(* IEC 61131-3 sources: codesys-conveyor-sorting/src, 4 files *)

(* ---- E_ConveyorState.st ---- *)
// DUT: E_ConveyorState
// States of the conveyor sorting station.
// Numbering in steps of 10 leaves room for new states later.

{attribute 'qualified_only'}
{attribute 'strict'}
TYPE E_ConveyorState :
(
    IDLE        := 0,   // Conveyor stopped, waiting for start
    RUNNING     := 10,  // Conveyor running, waiting for a part at the infeed
    CLASSIFYING := 20,  // Part detected, reading classification sensors
    TRANSPORT   := 30,  // Part travelling to the diverter, jam timer active
    DIVERTING   := 40,  // Diverter pulse active, part counted at the end
    FAULT       := 90,  // Jam detected, conveyor stopped, waiting for reset
    ESTOP       := 99   // E-stop active, all outputs off
);
END_TYPE

(* ---- E_PartType.st ---- *)
// DUT: E_PartType
// Result of the part classification at the infeed.

{attribute 'qualified_only'}
{attribute 'strict'}
TYPE E_PartType :
(
    NONE   := 0,  // No part being tracked
    TYPE_A := 1,  // Goes to bin A
    TYPE_B := 2,  // Goes to bin B
    REJECT := 3   // Unknown part (both or neither sensor), runs to reject bin
);
END_TYPE

(* ---- GVL_IO.st ---- *)
// GVL: GVL_IO
// Inputs and outputs of the sorting station.
// In this project they are driven by the CODESYS visualisation (simulation).
// On real hardware each variable would be mapped to a physical channel
// in the I/O configuration of the fieldbus device.

{attribute 'qualified_only'}
VAR_GLOBAL
    // ---- Digital inputs ----
    xStartPB         : BOOL;          // Start push button (TRUE = pressed)
    xStopPB          : BOOL;          // Stop push button (TRUE = pressed)
    xResetPB         : BOOL;          // Fault reset push button
    xEStopOK         : BOOL := TRUE;  // E-stop circuit healthy (NC contact, TRUE = OK)
    xPartAtEntry     : BOOL;          // Photo sensor at the infeed
    xSensorTypeA     : BOOL;          // Classification sensor, TRUE = type A
    xSensorTypeB     : BOOL;          // Classification sensor, TRUE = type B
    xPartAtDiverter  : BOOL;          // Photo sensor at the diverter position

    // ---- Digital outputs ----
    xConveyorRun     : BOOL;          // Conveyor motor contactor / VFD run command
    xDiverterA       : BOOL;          // Pneumatic diverter to bin A
    xDiverterB       : BOOL;          // Pneumatic diverter to bin B
    xLampRunning     : BOOL;          // Green lamp
    xLampFault       : BOOL;          // Red lamp (steady = jam, blinking = E-stop)
END_VAR

(* ---- PLC_PRG.st ---- *)
// =====================================================================
// POU: PLC_PRG (Program, Structured Text)
// Conveyor sorting station - main state machine
//
// Sequence: IDLE -> RUNNING -> CLASSIFYING -> TRANSPORT -> DIVERTING -> RUNNING
// Faults:   jam timeout -> FAULT, E-stop -> ESTOP (both need reset, then start)
//
// Note: the real E-stop is a hardwired safety circuit. The PLC only
// monitors it (xEStopOK) to stop the sequence and show the state.
// =====================================================================

// ---------------- DECLARATION (top pane in CODESYS) ----------------
PROGRAM PLC_PRG
VAR
    eState            : E_ConveyorState := E_ConveyorState.IDLE;
    ePartType         : E_PartType := E_PartType.NONE;
    xStopRequest      : BOOL;     // Stop pressed: finish the current part, then stop

    // Edge detection
    rtStart           : R_TRIG;
    rtReset           : R_TRIG;
    rtPartAtEntry     : R_TRIG;
    rtPartAtDiverter  : R_TRIG;

    // Timers
    tonJam            : TON;      // Part must reach the diverter within T_JAM_TIMEOUT
    tonDivert         : TON;      // Length of the diverter pulse
    tonBlink          : TON;      // Blink clock for the fault lamp
    xBlink            : BOOL;

    // Production counters (read later by the OPC UA data logger)
    udiCountA         : UDINT;
    udiCountB         : UDINT;
    udiCountReject    : UDINT;
    udiCountJams      : UDINT;
END_VAR
VAR CONSTANT
    T_JAM_TIMEOUT     : TIME := T#5S;
    T_DIVERT_PULSE    : TIME := T#500MS;
    T_BLINK           : TIME := T#500MS;
END_VAR

// ---------------- IMPLEMENTATION (bottom pane in CODESYS) ----------------

// ---- Edge detection ----
rtStart(CLK := GVL_IO.xStartPB);
rtReset(CLK := GVL_IO.xResetPB);
rtPartAtEntry(CLK := GVL_IO.xPartAtEntry);
rtPartAtDiverter(CLK := GVL_IO.xPartAtDiverter);

// ---- Timers (called every scan, outside the CASE) ----
tonJam(IN := (eState = E_ConveyorState.TRANSPORT), PT := T_JAM_TIMEOUT);
tonDivert(IN := (eState = E_ConveyorState.DIVERTING), PT := T_DIVERT_PULSE);
tonBlink(IN := NOT tonBlink.Q, PT := T_BLINK);
IF tonBlink.Q THEN
    xBlink := NOT xBlink;
END_IF

// ---- E-stop has priority over every state ----
IF NOT GVL_IO.xEStopOK THEN
    eState := E_ConveyorState.ESTOP;
END_IF

// ---- Stop request is latched and handled by the states ----
IF GVL_IO.xStopPB THEN
    xStopRequest := TRUE;
END_IF

// ---- State machine ----
CASE eState OF

    E_ConveyorState.IDLE:
        xStopRequest := FALSE;
        ePartType := E_PartType.NONE;
        IF rtStart.Q AND GVL_IO.xEStopOK THEN
            eState := E_ConveyorState.RUNNING;
        END_IF

    E_ConveyorState.RUNNING:
        IF xStopRequest THEN
            eState := E_ConveyorState.IDLE;
        ELSIF rtPartAtEntry.Q THEN
            eState := E_ConveyorState.CLASSIFYING;
        END_IF

    E_ConveyorState.CLASSIFYING:
        // Exactly one sensor must be active, otherwise the part is rejected
        IF GVL_IO.xSensorTypeA AND NOT GVL_IO.xSensorTypeB THEN
            ePartType := E_PartType.TYPE_A;
        ELSIF GVL_IO.xSensorTypeB AND NOT GVL_IO.xSensorTypeA THEN
            ePartType := E_PartType.TYPE_B;
        ELSE
            ePartType := E_PartType.REJECT;
        END_IF
        eState := E_ConveyorState.TRANSPORT;

    E_ConveyorState.TRANSPORT:
        IF rtPartAtDiverter.Q THEN
            eState := E_ConveyorState.DIVERTING;
        ELSIF tonJam.Q THEN
            udiCountJams := udiCountJams + 1;
            eState := E_ConveyorState.FAULT;
        END_IF

    E_ConveyorState.DIVERTING:
        IF tonDivert.Q THEN
            CASE ePartType OF
                E_PartType.TYPE_A:
                    udiCountA := udiCountA + 1;
                E_PartType.TYPE_B:
                    udiCountB := udiCountB + 1;
            ELSE
                udiCountReject := udiCountReject + 1;
            END_CASE
            ePartType := E_PartType.NONE;

            IF xStopRequest THEN
                eState := E_ConveyorState.IDLE;
            ELSE
                eState := E_ConveyorState.RUNNING;
            END_IF
        END_IF

    E_ConveyorState.FAULT:
        // Operator clears the jam, then presses reset
        IF rtReset.Q THEN
            eState := E_ConveyorState.IDLE;
        END_IF

    E_ConveyorState.ESTOP:
        // E-stop must be released AND reset pressed; no automatic restart
        IF GVL_IO.xEStopOK AND rtReset.Q THEN
            eState := E_ConveyorState.IDLE;
        END_IF

END_CASE

// ---- Outputs: written in one place only ----
GVL_IO.xConveyorRun := (eState = E_ConveyorState.RUNNING)
                    OR (eState = E_ConveyorState.CLASSIFYING)
                    OR (eState = E_ConveyorState.TRANSPORT)
                    OR (eState = E_ConveyorState.DIVERTING);

GVL_IO.xDiverterA   := (eState = E_ConveyorState.DIVERTING) AND (ePartType = E_PartType.TYPE_A);
GVL_IO.xDiverterB   := (eState = E_ConveyorState.DIVERTING) AND (ePartType = E_PartType.TYPE_B);

GVL_IO.xLampRunning := GVL_IO.xConveyorRun;
GVL_IO.xLampFault   := (eState = E_ConveyorState.FAULT)
                    OR ((eState = E_ConveyorState.ESTOP) AND xBlink);
